// TIA Portal V21 export
// export: Created 2026-11-11T00:49:05.9908593Z, ExportSetting WithDefaults, DisplayName Totally Integrated Automation Portal, DisplayVersion V21 Update 3, DisplayName STEP 7 Professional, DisplayVersion V21 Update 3, DisplayName STEP 7 Safety, DisplayVersion V21, DisplayName Tech WebApplication, DisplayVersion V21, DisplayName WinCC Basic/Comfort/Advanced, DisplayVersion V21 Update 3, DisplayName WinCC Unified, DisplayVersion V21 Update 3
FUNCTION_BLOCK "FX_Lad_pt001"   // FB250, LAD
{ S7_Optimized_Access := 'TRUE' }
VERSION : 0.1
// stored: AutoNumber true, IsIECCheckEnabled false, IsRetainMemResEnabled false, MemoryReserve 100, SetENOAutomatically false, UDAEnableTagReadback false
   VAR_INPUT
      "a" : Bool;
      "b" : Bool;
      c : Bool;
      ia : Int;
      ib : Int;
      ic : Int;
      da : DInt;
      db : DInt;
      ra : Real;
      rb : Real;
      wa : Word;
      wb : Word;
      dwa : DWord;
      ba : Byte;
      ta : Time;
      tb : Time;
      s1 : String;
      s2 : String;
   END_VAR
   VAR_OUTPUT
      q : Bool;
      q2 : Bool;
      io : Int;
      io2 : Int;
      dout : DInt;
      rout : Real;
      wout : Word;
      dwout : DWord;
      bout : Byte;
      tout : Time;
      sout : String;
   END_VAR
   VAR_IN_OUT
      p_req : Bool;
      p_port : PORT;
      p_protocol : UInt;
      p_baud : UInt;
      p_parity : UInt;
      p_databits : UInt;
      p_stopbits : UInt;
      p_flowctrl : UInt;
      p_xonchar : Char;
      p_xoffchar : Char;
      p_waittime : UInt;
      p_done : Bool;
      p_error : Bool;
      p_status : Word;
      x_usint : USInt;
      arr : Array[0..9] of Int;
      barr : Array[0..7] of Bool;
      iinout : Int;
   END_VAR
   VAR
      inst : Port_Config;
      ton1 { S7_SetPoint := 'True'} : TON_TIME;
      tof1 { S7_SetPoint := 'True'} : TOF_TIME;
      tp1 { S7_SetPoint := 'True'} : TP_TIME;
      tonr1 { S7_SetPoint := 'True'} : TONR_TIME;
      ctu1 { S7_SetPoint := 'True'} : CTU_INT;
      ctd1 { S7_SetPoint := 'True'} : CTD_INT;
      ctud1 { S7_SetPoint := 'True'} : CTUD_INT;
      rtrig1 { S7_SetPoint := 'True'} : R_TRIG;
      ftrig1 { S7_SetPoint := 'True'} : F_TRIG;
      edge1 : Bool;
      edge2 : Bool;
      stat1 : Bool;
      stat2 : Bool;
      stati : Int;
   END_VAR
   VAR_TEMP
      t1 : Bool;
      t2 : Bool;
      ti : Int;
      td : DInt;
      tr : Real;
      tw : Word;
      tt : Time;
      var1 : Variant;
   END_VAR
BEGIN

REGION Network 1: ---| |--- - Normally open contact
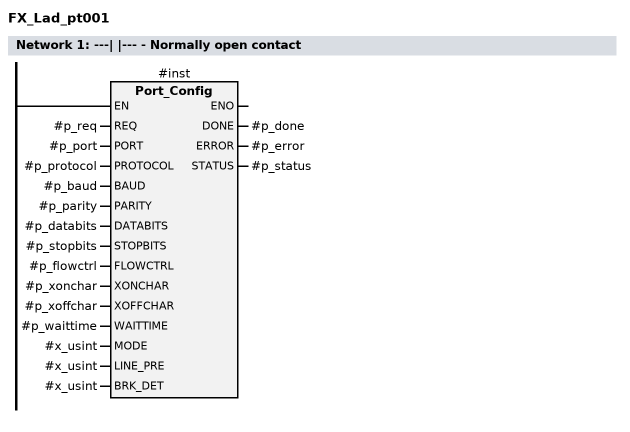
   RUNG wire#powerrail
      #inst.Port_Config(REQ := #p_req, PORT := #p_port, PROTOCOL := #p_protocol, BAUD := #p_baud, PARITY := #p_parity, DATABITS := #p_databits, STOPBITS := #p_stopbits, FLOWCTRL := #p_flowctrl, XONCHAR := #p_xonchar, XOFFCHAR := #p_xoffchar, WAITTIME := #p_waittime, DONE => #p_done, ERROR => #p_error, STATUS => #p_status, MODE := #x_usint, LINE_PRE := #x_usint, BRK_DET := #x_usint)
   END_RUNG
   // the same network as SCL:
   #inst(REQ := #p_req,   // Port_Config
         PORT := #p_port,
         PROTOCOL := #p_protocol,
         BAUD := #p_baud,
         PARITY := #p_parity,
         DATABITS := #p_databits,
         STOPBITS := #p_stopbits,
         FLOWCTRL := #p_flowctrl,
         XONCHAR := #p_xonchar,
         XOFFCHAR := #p_xoffchar,
         WAITTIME := #p_waittime,
         MODE := #x_usint,
         LINE_PRE := #x_usint,
         BRK_DET := #x_usint,
         DONE => #p_done,
         ERROR => #p_error,
         STATUS => #p_status);
END_REGION
END_FUNCTION_BLOCK
